# B&R Automation Studio project lab1
Automation Studio 4.5.2.102

## Configuration sim

CPU 4PP065.0571-P74, AutomationRuntime D4.52, Build 4.1.2, Vc V4.52.0

### Task classes (Cpu.sw)
```
Cyclic#4:
  Program <- Program.prg
Binaries: udbdef, TCData, iomap, ashwac, Role, sysconf, arconfig, asfw, User, ashwd
Libraries: Library
```

### Hardware
```
4PP065_0571_P74 : 4PP065.0571-P74 v1.1.2.0
  Connector IF5:
    ActivateDevice = 1
  ConfigurationID = labBR
  Simulation = 1
```

- Physical/sim/4PP065_0571_P74/IoMap.iom: same as Physical/sim/4PP065_0571_P74/Cpu.per
- Physical/sim/4PP065_0571_P74/PvMap.vvm: same as Physical/sim/4PP065_0571_P74/Cpu.per
## Logical view

Binary libraries used (declarations not repeated): operator, runtime, astime, AsIecCon

### Package Logical/Libraries - Global libraries

### Library Logical/Libraries/Library (ANSIC)

#### Library.fun - Exported functions and function blocks
```iecst
{REDUND_ERROR} {REDUND_UNREPLICABLE} FUNCTION_BLOCK FB_Motor (*TODO: Add your comment here*) (*$GROUP=User,$CAT=User,$GROUPICON=User.png,$CATICON=User.png*)
	VAR_INPUT
		u : {REDUND_UNREPLICABLE} REAL;
	END_VAR
	VAR_OUTPUT
		w : {REDUND_UNREPLICABLE} REAL;
		phi : {REDUND_UNREPLICABLE} REAL;
	END_VAR
	VAR
		integrator2 : {REDUND_UNREPLICABLE} FB_Integrator;
		integrator : {REDUND_UNREPLICABLE} FB_Integrator;
		Tm : {REDUND_UNREPLICABLE} REAL;
		ke : {REDUND_UNREPLICABLE} REAL;
		dt : {REDUND_UNREPLICABLE} REAL;
	END_VAR
END_FUNCTION_BLOCK

{REDUND_ERROR} FUNCTION_BLOCK FB_Integrator (*TODO: Add your comment here*) (*$GROUP=User,$CAT=User,$GROUPICON=User.png,$CATICON=User.png*)
	VAR_INPUT
		in : {REDUND_UNREPLICABLE} REAL;
	END_VAR
	VAR_OUTPUT
		out : {REDUND_UNREPLICABLE} REAL;
	END_VAR
	VAR
		dt : {REDUND_UNREPLICABLE} REAL;
		star : REAL;
	END_VAR
END_FUNCTION_BLOCK

{REDUND_ERROR} {REDUND_UNREPLICABLE} FUNCTION_BLOCK FB_Regulator (*TODO: Add your comment here*) (*$GROUP=User,$CAT=User,$GROUPICON=User.png,$CATICON=User.png*)
	VAR_INPUT
		e : {REDUND_UNREPLICABLE} REAL;
	END_VAR
	VAR_OUTPUT
		u : {REDUND_UNREPLICABLE} REAL;
	END_VAR
	VAR
		k_p : {REDUND_UNREPLICABLE} REAL;
		k_i : {REDUND_UNREPLICABLE} REAL;
		integrator : {REDUND_UNREPLICABLE} FB_Integrator;
		iyOld : {REDUND_UNREPLICABLE} REAL;
		max_abs_value : {REDUND_UNREPLICABLE} REAL;
		dt : {REDUND_UNREPLICABLE} REAL;
	END_VAR
END_FUNCTION_BLOCK
```

#### FB_Motor.c
```c
#include <bur/plctypes.h>
#ifdef __cplusplus
	extern "C"
	{
#endif
	#include "Library.h"
#ifdef __cplusplus
	};
#endif
/* TODO: Add your comment here */
void FB_Motor(struct FB_Motor* inst)
{
    REAL U = inst->u / inst->ke;
    REAL wich = (U-inst->w) /inst->Tm;
    inst->integrator.in = wich;
    FB_Integrator(&inst->integrator);
    inst->w = inst->integrator.out;
    inst->integrator2.in = inst->w;
    FB_Integrator(&inst->integrator2);
    inst->phi = inst->integrator2.out;
}
```

#### FB_Integrator.c
```c
#include <bur/plctypes.h>
#ifdef __cplusplus
	extern "C"
	{
#endif
	#include "Library.h"
#ifdef __cplusplus
	};
#endif
/* TODO: Add your comment here */
void FB_Integrator(struct FB_Integrator* inst)
{
    inst->dt = 0.01;
    inst->out = inst->out + inst->in * inst->dt;
    inst->star = inst->out;
}
```

#### FB_Regulator.c
```c
#include <bur/plctypes.h>
#ifdef __cplusplus
	extern "C"
	{
#endif
	#include "Library.h"
#ifdef __cplusplus
	};
#endif
/* TODO: Add your comment here */
void FB_Regulator(struct FB_Regulator* inst)
{
    REAL p1 = inst->e * inst->k_p;

    REAL p2 = inst->e * inst->k_i;

    inst->integrator.in = p2 + inst->iyOld;
    FB_Integrator(&inst->integrator);
    REAL r = inst->integrator.out;
    REAL p3 = p1 + r;
    REAL pered = p3;
    REAL lim;
    if (pered > inst->max_abs_value)   lim=inst->max_abs_value;
    else if (pered < -inst->max_abs_value)   lim=-inst->max_abs_value;
    else lim = pered;
    REAL correction = lim - pered;
    inst->iyOld = r+ correction;
    inst->u = lim;
}
```

### Program Logical/Program (ANSIC)

#### Cyclic.c - Cyclic code
```c
#include <bur/plctypes.h>

#ifdef _DEFAULT_INCLUDES
	#include <AsDefault.h>
#endif

void _CYCLIC ProgramCyclic(void)
{

    counter++;
    if ((counter >= 300) && (counter <= 800))
        speed = 100;
    else
        speed = 0;

    // áåç ðåã
    fb_motor2.u = speed * fb_motor2.ke;
    FB_Motor(&fb_motor2);
    // ñ ðåã
    fb_regulator.e = speed  - fb_motor.w;
    FB_Regulator(&fb_regulator);
    fb_motor.u = fb_regulator.u;
    FB_Motor(&fb_motor);

}
```

#### Init.c - Initialization code
```c
#include <bur/plctypes.h>

#ifdef _DEFAULT_INCLUDES
	#include <AsDefault.h>
#endif

void _INIT ProgramInit(void)
{
     fb_motor.Tm = 0.06;
     fb_motor.ke = 27.0/145.0;
     fb_motor.dt = 0.01;

    fb_motor2.Tm = 0.06;
    fb_motor2.ke = 27.0/145.0;
    fb_motor2.dt = 0.01;

    fb_regulator.k_i = fb_motor.ke / 0.03;
    fb_regulator.k_p = (fb_motor.ke * fb_motor.Tm) / 0.03;
    fb_regulator.max_abs_value = 27;
    fb_regulator.dt = 0.01;
    fb_regulator.iyOld = 0;

    speed = 0;
    enable = 1;
    counter = 0;
}
```

#### Exit.c - Exit code
```c
#include <bur/plctypes.h>

#ifdef _DEFAULT_INCLUDES
	#include <AsDefault.h>
#endif

void _EXIT ProgramExit(void)
{

}
```

#### Variables.var - Local variables
```iecst
VAR
	fb_regulator : FB_Regulator;
	fb_motor2 : FB_Motor;
	fb_motor : FB_Motor;
	speed : REAL;
	counter : UINT;
	enable : BOOL;
END_VAR
```
